TYPE TwinSafeIn_PlcOut :
STRUCT
	RUN			: BOOL;
	ErrACK		: BOOL;
	//Restart		: BOOL; //Restart TwinSAFE
END_STRUCT
END_TYPE

(* stored: Version 1.1.0.1, ProductVersion 3.1.4024.13
   DUT TwinSafeIn_PlcOut: Id {21e586ed-5092-41e6-9ebf-c0ef0cc442c5} *)
